Fanuc KAREL source: kt00446.KL

-- PROVISIONAL review KL for V770-1; original PC SHA256 0d152f5f1e43dcc17a19170f3e3c1e8106bbf10223f531522ce85671e31c2b75
-- Incomplete behavior may be omitted. Consult companion uncertainty JSON. Do not deploy.
PROGRAM KT00446
%NOLOCKGROUP
VAR
  S1 : STRING[80]
  S2 : STRING[80]
  OUT : BOOLEAN
BEGIN
  -- UNRESOLVED_PC offsets 5-14; opcodes 3F,75
  -- UNRESOLVED_PC offsets 19-28; opcodes 3F,75
  -- UNRESOLVED_PC offsets 33-42; opcodes 3F,75
  -- UNRESOLVED_PC offsets 47-56; opcodes 3F,75
  -- UNRESOLVED_PC offsets 61-80; opcodes 73,73,88,23
  -- UNRESOLVED_PC offsets 85-89; opcodes 7F
END KT00446
